(* IEC 61131-3 sources: 2026_Projet_YGO_ExcavatriceDragage/CODE/J_SUPERVISION/_TYPES/2_TRANSLATION, 17 files *)

(* ---- E_TranslationTraceBlockReason.st ---- *)
(* =======================================================================
   🎯 E_TranslationTraceBlockReason — Cause de blocage priorisée translation M3
   ───────────────────────────────────────────────────────────────
   🎯 Rôle : Ordre de priorité de la cause de blocage de la translation M3,
      calculé en PRG_05_Translation et publié via Data.TranslationTrace.
      L'ordre de l'enum EST l'ordre de priorité (valeur croissante = priorité
      décroissante) : la cause la plus grave gagne (PowerCutOff > … > NONE).
   📤 Producteur unique : PRG_05_Translation.
   📥 Consommateur : FB_TroubleshootingView (recopie → GVL_Troubleshooting.S_TraceTranslation).
   🔒 Lecture seule — aucune action de conduite n'en dépend.
   📄 Doc métier : DOC/AF/AF_Partie-14_Fonction_Troubleshooting/FB_TroubleshootingView_v1.2.md
   ======================================================================= *)
{attribute 'qualified_only'}
TYPE E_TranslationTraceBlockReason :
(
    NONE              := 0,   // ✅ Aucun blocage — permis de mouvement effectif
    POWER_CUTOFF      := 1,   // 🧨 Coupure puissance amont (instSafetyTranslationM3.PowerCutOff) — priorité max
    SAFESTOP          := 2,   // 🟧 SafeStop effectif (InputModule OR safety M3)
    SAFETY_FAULT      := 3,   // 🛡️ Défaut safety M3 latched (FB_Safety_Translation.Fault.Error)
    HEIGHT_INTERLOCK  := 4,   // 🚧 Interlock hauteur M1/M2 actif (risque collision)
    DRIVE_UNAVAILABLE := 5,   // 📡 Variateur AC600 injoignable / non opérationnel
    FINAL_INTERLOCK   := 6,   // 🛑 Barrière finale en défaut (frein / redémarrage)
    FAULT             := 7    // ❌ Défaut mouvement M3 latched (FB_Translation.Fault.Error)
);
END_TYPE

(* ---- ST_BypassTranslation.st ---- *)
(* ═══════════════════════════════════════════════════════════════
   ST_BypassTranslation — Bypass maintenance dédiés à Translation M3
   ───────────────────────────────────────────────────────────────
   🔒 Doctrine : actionnable UNIQUEMENT en MAINT_N2, RETAIN, jamais masque
      les autres défauts du même bloc (voir REGISTRE_ACTIONS_Bypass_v1.0 (archive)).
   ═══════════════════════════════════════════════════════════════ *)
TYPE ST_BypassTranslation :
STRUCT
    (* 📡 1. Communication & Systèmes auxiliaires *)
    OperatorComm      : BOOL; (* 📡 Bypass communication esclave CANopen Joystick / heartbeat IHM *)
    DriveComm         : BOOL; (* 📡 Bypass diagnostic esclave EtherCAT AC600 (variateur) *)
    ContactorFeedback : BOOL; (* 🔌 Bypass feedbacks contacteur de frein *)
    PhaseRotation     : BOOL; (* ⚡ Bypass défaut rotation de phases (commun machine) *)
    BrakeThermal      : BOOL; (* 🌡️ Bypass surchauffe thermique frein (commun machine) *)

    (* 🚧 2. Limites physiques et Positionnement *)
    LimitSwitch       : BOOL; (* 🚧 Bypass fins de course physiques avant/arrière *)
    SensorIncoherent  : BOOL; (* 🧭 Bypass incohérence mot capteurs de position *)
    MinHeight         : BOOL; (* : Bypass interlock hauteur mini M1/M2 requise pour translation *)

    (* ⚙️ 3. Sécurité Mécanique (Méca A-B) *)
    MecaA             : BOOL; (* 🔄 Bypass Méca A : mouvement non commandé à l'arrêt *)
    MecaB             : BOOL; (* 🛑 Bypass Méca B : absence confirmation arrêt (frein/contacteurs) *)

    (* 🛡️ 4. Hiérarchie & Restauration *)
    Safety            : BOOL; (* 🛡️ Bypass groupé : tous les bits qui provoquent un PowerCutOff *)
    Process           : BOOL; (* ⚙️ Bypass groupé : tous les bits qui provoquent un SafeStop *)
    Global            : BOOL; (* 🌐 Bypass Global : ignore toutes les sécurités de cet axe *)
    // Flag restauration boot dédié (défaut FALSE non ambigu, contrairement à une valeur métier)
    Initialized       : BOOL := FALSE; (* 🚦 TRUE = bypass restauré depuis GVL_BypassRetain ce boot *)
END_STRUCT
END_TYPE

(* ---- ST_Chain_Translation_Control.st ---- *)
TYPE ST_Chain_Translation_Control :
STRUCT
    Idx401_MotionAllowed         : BOOL; // 1 = Mouvement Translation Autorisé | 0 = Bloqué
    Idx402_SetpointFreq_Hz       : REAL; // [Hz] Consigne Fréquence Calculée
    Idx403_DriveControlWord      : WORD; // Mot de Commande Calculé Variateur AC600
    Idx404_FinalInterlockState   : E_State; // 🛡️ État frontière
    Idx405_FinalInterlockReason  : E_TranslationFinalInterlockReason; // 🛡️ Cause mémorisée
    Idx406_BrakeCommandOpenConfirmed : BOOL; // 🔌 Contacteur/bobine, pas frein mécanique
    Idx407_BrakeTimeoutElapsed   : TIME; // ⏱️ Watchdog 500ms écoulé
END_STRUCT
END_TYPE

(* ---- ST_Chain_Translation_Demandes.st ---- *)
TYPE ST_Chain_Translation_Demandes :
STRUCT
    Idx201_JoyXRaw_ANA           : INT;  // [pts] Bruts Joystick Axe X
    Idx202_JoyXScaled_Pct        : REAL; // [%] Consigne Joystick Axe X (-100% à +100%)
    Idx203_HmiCmd_BtnTremie : BOOL; // 1 = Bouton vers Trémie IHM | 0 = Relâché (ex-Idx203_HmiCmd_BtnFwd)
    Idx204_HmiCmd_BtnMaintenance : BOOL; // 1 = Bouton vers Maintenance IHM | 0 = Relâché (ex-Idx204_HmiCmd_BtnRev)
    Idx205_HmiTargetPosition     : INT;  // Cible Sélectionnée IHM (1=Trémie, 2=P2, 3=P1)
    Idx206_CycleTargetPosition   : INT;  // Cible Sélectionnée par le Cycle Auto
    Idx207_ModeActive            : E_Mode;// Mode courant (MANU_N1, AUTO_N1...)
    Idx208_BypassNetworkActive   : BOOL; // 0 = Comm Variateur OK | 1 = Bypass Réseau Actif ⚠️
    Idx209_ArbitratedSpeed_Pct   : REAL; // [%] Consigne finale Vitesse Translation
END_STRUCT
END_TYPE

(* ---- ST_Chain_Translation_Inputs.st ---- *)
TYPE ST_Chain_Translation_Inputs :
STRUCT
    Idx101_PosTremie_DI          : BOOL; // 1 = Position Trémie Atteinte | 0 = Absent
    Idx102_PosPV_DI              : BOOL; // 1 = Zone Ralentissement PV Atteinte | 0 = Absent
    Idx103_PosP2_DI              : BOOL; // 1 = Position Fosse P2 Atteinte | 0 = Absent
    Idx104_PosP1_DI              : BOOL; // 1 = Position Fosse P1 Atteinte | 0 = Absent
    Idx105_PosMaintenance_DI     : BOOL; // 1 = Position Service Maintenance Atteinte | 0 = Absent
    Idx106_DriveActualFreq_Hz    : REAL; // [Hz] Fréquence Réelle Mesurée Variateur
    Idx107_DriveStatusWord       : WORD; // Mot d'état Brut Variateur AC600
    Idx108_BrakeApplied          : BOOL; // TRUE = frein SERRÉ (NOT BrakeFeedback — IHM garde le sens serré)
    Idx109_DriveThermalOk        : BOOL; // TRUE = thermique moteur/variateur AC600 OK (diagnostic seul)
END_STRUCT
END_TYPE

(* ---- ST_Chain_Translation_Outputs.st ---- *)
TYPE ST_Chain_Translation_Outputs :
STRUCT
    Idx501_CmdDriveControlWord   : WORD; // Mot de Commande Transmis EtherCAT AC600
    Idx502_CmdDriveFreq_Hz       : UINT; // [0.01Hz] Consigne Fréquence Transmise EtherCAT
    Idx503_CmdBrakeRelease_RQ    : BOOL; // 1 = Bobine Frein Translation Alimentée (Ouvert)
END_STRUCT
END_TYPE

(* ---- ST_Chain_Translation_Safety.st ---- *)
TYPE ST_Chain_Translation_Safety :
STRUCT
    Idx301_EmergencyChainClosed  : BOOL; // 1 = Boucle Urgence OK | 0 = Arrêt d'Urgence Appuyé
    Idx302_SafeStopActive        : BOOL; // 0 = Sain (Autorisé) | 1 = Arrêt Rapide Translation
    Idx303_PowerCutOffActive     : BOOL; // 0 = Puissance OK | 1 = Coupure Puissance
    Idx304_LimitSwitchTremieActive  : BOOL; // 0 = Sain | 1 = Fin de Course Extrême Trémie (ex-Idx304_LimitSwitchFwdActive)
    Idx305_LimitSwitchMaintenanceActive : BOOL; // 0 = Sain | 1 = Fin de Course Extrême Maintenance (ex-Idx305_LimitSwitchRevActive)
    Idx306_BypassLimitSwitch     : BOOL; // 0 = Fins de course actives | 1 = Shuntés IHM ⚠️
    Idx307_PositionDecoderIncoherent: BOOL; // 0 = Décodage 5 Capteurs OK | 1 = Incohérence Position
    Idx308_HeightInterlockBlocking: BOOL; // : 0 = M1 ET M2 ≥ hauteur mini (ou bypass) | 1 = Translation bloquée (risque collision)
    (* Défauts safety déchiffrés (bits ErrorId) — visibles individuellement à l'IHM *)
    Idx309_ErrorOperatorComm : BOOL; // bit0 Perte communication opérateur (joystick CAN / heartbeat IHM)
    Idx310_ErrorDriveComm    : BOOL; // bit1 Perte communication EtherCAT variateur
    Idx311_ErrorPhaseRotation: BOOL; // bit2 Mauvaise rotation de phases
    Idx312_ErrorBrakeThermal : BOOL; // bit3 Surchauffe thermique frein commun
    Idx313_ErrorMecaB        : BOOL; // bit4 Absence confirmation arrêt
    Idx314_ErrorMecaA        : BOOL; // bit5 Mouvement non commandé
    Idx315_ErrorLimitSwitch  : BOOL; // bit6 Limite extrême atteinte
    Idx316_ErrorSensorIncoherent: BOOL; // bit7 Mot capteurs position incohérent
    Idx317_ErrorId           : WORD; // Masque brut complet (latch cause) — source d'arbitrage PowerCutOff
    (* Permis directionnels M3 (source unique : FB_Safety_Translation) — TRUE = autorisé, fail-safe *)
    Idx318_EffectivePermitM3_Tremie      : BOOL; // 1 = Translation vers Trémie autorisée | 0 = SENS TRÉMIE BLOQUÉ
    Idx319_EffectivePermitM3_Maintenance : BOOL; // 1 = Translation vers Maintenance/P1 autorisée | 0 = SENS MAINTENANCE BLOQUÉ
END_STRUCT
END_TYPE

(* ---- ST_ChainTranslation.st ---- *)
TYPE ST_ChainTranslation :
STRUCT
    Inputs_100    : ST_Chain_Translation_Inputs;
    Demandes_200  : ST_Chain_Translation_Demandes;
    Safety_300    : ST_Chain_Translation_Safety;
    Control_400   : ST_Chain_Translation_Control;
    Outputs_500   : ST_Chain_Translation_Outputs;
END_STRUCT
END_TYPE

(* ---- ST_HwTranslation.st ---- *)
(* ═══════════════════════════════════════════════════════════════
   🏗️ ST_HwTranslation — Image matérielle brute des entrées Translation M3
   ───────────────────────────────────────────────────────────────
   🎨 Regroupe les signaux physiques d'entrée bruts de la translation M3 (AC600).
   ═══════════════════════════════════════════════════════════════ *)
TYPE ST_HwTranslation :
STRUCT
    M3_PosTremie_DI      : BOOL;         (* Capteur position trémie *)
    M3_PosPV_DI          : BOOL;         (* Capteur position point de vitesse (pré-ralentissement) *)
    M3_PosPVP2_DI        : BOOL;         (* Capteur position P2 / petite vitesse avant P1 *)
    M3_PosP1_DI          : BOOL;         (* Capteur position P1 *)
    M3_PosMaintenance_DI : BOOL;         (* Capteur position maintenance *)
    M3_BrakeIsOpen_DI    : BOOL;         (* Retour frein M3 (1 = ouvert) *)
    M3_ThermalOK_DI      : BOOL;         (* Retour disjoncteur thermique moteur/variateur AC600 (1 = OK) — diagnostic seul, l'AC600 se protège lui-même *)
    M3_StatusWord        : WORD;         (* Status word variateur AC600 *)
    M3_ActualFrequencyHz : UINT;         (* Fréquence réelle variateur AC600 (x100) *)
    AC600_DeviceState    : DEVICE_STATE; (* État device AC600 (GetDeviceState) *)
END_STRUCT
END_TYPE

(* ---- ST_SafetyTranslation.st ---- *)
(* ═══════════════════════════════════════════════════════════════
   🛡️ ST_SafetyTranslation — Diagnostics de sécurité pour la Translation M3
   ───────────────────────────────────────────────────────────────
   🎨 Destiné à l'affichage des défauts de sécurité du translation.
   ═══════════════════════════════════════════════════════════════ *)
TYPE ST_SafetyTranslation :
STRUCT
    Error             : BOOL;    (* 🛡️ Bloc sécurité (Safety) en défaut *)
    ErrorId           : WORD;    (* ❌ Code bitfield du défaut de sécurité (vue LIVE) *)
    LatchedId         : WORD;    (* 🕘 Vue LATCHÉE : ErrorId figé au défaut, effacé au Reset (marqueur [HISTO]) *)
    ErrorOperatorComm : BOOL;    (* 🎮 Perte communication opérateur : joystick CAN ou heartbeat IHM (bit0) *)
    ErrorDriveComm    : BOOL;    (* 📡 Perte communication EtherCAT variateur (bit1) *)
    ErrorPhaseRotation: BOOL;    (* ⚡ Mauvaise rotation de phases électriques (bit2) *)
    ErrorBrakeThermal : BOOL;    (* 🌡️ Surchauffe thermique frein commun (bit3) *)
    ErrorMecaB        : BOOL;    (* 🛑 Absence confirmation arrêt (Méca B - bit4) *)
    ErrorMecaA        : BOOL;    (* 🔄 Mouvement non commandé (Méca A - bit5) *)
    ErrorLimitSwitch  : BOOL;    (* 🚧 Limite extrême Translation atteinte (bit6) *)
    ErrorSensorIncoherent : BOOL; (* 🧭 Mot capteurs M3 incohérent (bit7) *)
    SafeStop          : BOOL;    (* 🛡️ Décélération de sécurité demandée *)
    PowerCutOff       : BOOL;    (* 🧨 Coupure puissance demandée *)
    EffectivePermitM3_Tremie      : BOOL;    (* 🟢 Permis canonique M3 vers Trémie, TRUE = autorisé *)
    EffectivePermitM3_Maintenance : BOOL;    (* 🟢 Permis canonique M3 vers Maintenance/P1, TRUE = autorisé *)
    BlockedBySafety   : BOOL;    (* 🚫 Synthèse globale : translation bloquée par la sécurité *)
    PowerCutOffSafety : BOOL;    (* 🧨 Synthèse sécurités critiques entraînant une coupure puissance *)
    SafeStopSafety    : BOOL;    (* 🛡️ Synthèse défauts entraînant un SafeStop / Rampe rapide *)
END_STRUCT
END_TYPE

(* ---- ST_TraceTranslation.st ---- *)
(* =======================================================================
   ↔️ ST_TraceTranslation — Trace de blocage terrain de la translation M3
   ───────────────────────────────────────────────────────────────
   🎯 Rôle : Publier au technicien « pourquoi la translation M3 ne bouge pas » :
      permis de mouvement effectif, interlock hauteur, source SafeStop/coupure
      et cause de blocage priorisée.
   📤 Producteur unique : PRG_05_Translation (Data.TranslationTrace).
   📥 Consommateur : FB_TroubleshootingView (pure recopie → GVL_Troubleshooting.S_TraceTranslation).
   🔒 Lecture seule — aucun calcul de commande n'en dépend.
   🕒 BlockReasonTimestamp : ms depuis démarrage PLC (TIME()), latched au dernier
      changement de BlockReason (1 scan, mémoire).
   📄 Doc métier : DOC/AF/AF_Partie-14_Fonction_Troubleshooting/FB_TroubleshootingView_v1.2.md
   ======================================================================= *)
TYPE ST_TraceTranslation :
STRUCT
    // Permis de mouvement effectif (agrégat diagnostic : toutes les barrières levées)
    MotionPermitEffective    : BOOL;   // 🟢 Translation réellement autorisée à se déplacer
    // Permis directionnels par sens (reflet exact des permis appliqués au mouvement M3)
    EffectivePermitM3_Tremie      : BOOL;   // 🟢 Permis canonique M3 vers Trémie (reflet lecture seule)
    EffectivePermitM3_Maintenance : BOOL;   // 🟢 Permis canonique M3 vers Maintenance/P1 (reflet lecture seule)
    TremieProcessBlockActive : BOOL;   // 🛑 Approche trémie interdite par process (trémie pleine / grille levée) — recul libre. Motif du permis trémie rouge.
    HeightInterlockBlocking  : BOOL;   // 🚧 Interlock hauteur M1/M2 actif (risque collision)

    // Source de blocage — pour distinguer l'origine
    SafeStopActive           : BOOL;   // 🟧 SafeStop effectif appliqué (M3_SafeStop_Aggregate)
    SafeStopSourceInput      : BOOL;   // 📥 SafeStop issu du module d'entrée (InputModuleFault)
    SafeStopSourceSafety     : BOOL;   // 🛡️ SafeStop issu de FB_Safety_Translation (défaut safety)
    PowerCutOffActive        : BOOL;   // 🧨 Coupure puissance amont active
    DriveOperational         : BOOL;   // 📡 Variateur AC600 opérationnel

    // Barrière finale (frein / redémarrage)
    FinalInterlockError      : BOOL;   // 🛑 Défaut barrière finale (frein / redémarrage)

    // Cause de blocage priorisée + horodatage
    BlockReason              : E_TranslationTraceBlockReason; // 🎯 Cause de blocage prioritaire (ordre de priorité croissant)
    BlockReasonTimestamp     : UDINT;  // 🕒 ms depuis démarrage PLC (TIME()) — dernier changement de BlockReason
END_STRUCT
END_TYPE

(* ---- ST_TranslationCfg.st ---- *)
(* ═══════════════════════════════════════════════════════════════
   ST_TranslationCfg — Configurations et paramètres réglables pour Translation M3
   ───────────────────────────────────────────────────────────────
   🎨 Destiné au paramétrage depuis l'IHM (RETAIN) — même patron que ST_WinchCfg.
   📄 Vitesses de ralentissement d'approche réglables depuis l'IHM (RETAIN), même patron que ST_WinchCfg.
   ═══════════════════════════════════════════════════════════════ *)
TYPE ST_TranslationCfg :
STRUCT
    CfgApproachSpeedTremie_Hz      : REAL := 20.0; (* 🐢 Vitesse réduite d'approche Trémie (Hz), déclenchée par capteur PV, Direction=1 — reglage nominal confirme operateur *)
    CfgApproachSpeedMaintenance_Hz : REAL := 20.0; (* 🐢 Vitesse réduite d'approche Maintenance (Hz), déclenchée par capteur P1, Direction=-1 — reglage nominal confirme operateur *)
    CfgApproachSpeedP1_Hz          : REAL := 20.0; (* 🐢 Vitesse réduite d'approche P1 (Hz), déclenchée par capteur P2, Direction=-1 — reglage nominal confirme operateur *)

    (* Flag restauration boot (défaut FALSE non ambigu) — même patron que ST_WinchCfg *)
    Initialized                    : BOOL := FALSE; (* 🚦 TRUE = config restaurée depuis GVL_PERSISTENT ce boot *)
END_STRUCT
END_TYPE

(* ---- ST_TranslationCmd.st ---- *)
(* ═══════════════════════════════════════════════════════════════
   🎮 ST_TranslationCmd — Commandes IHM pour la Translation M3
   ───────────────────────────────────────────────────────────────
   🎨 Destiné au pilotage de la translation M3 depuis l'IHM.
   📄 : Initialized protège SetFreq_Hz (seul réglage à survivre au reboot),
      sans pont générique pour ne jamais persister BtnTremie/BtnMaintenance.
   ═══════════════════════════════════════════════════════════════ *)
TYPE ST_TranslationCmd :
STRUCT
    SelPositioning     : BOOL;    (* 🎯 TRUE = positionneur sur SelTarget ; FALSE = jog libre *)
    SelTarget          : INT;     (* 🔢 Numéro de la cible de position sélectionnée *)
    BtnTremie         : BOOL;    (* ↔️ Requête marche vers Trémie (ex-BtnFwd), pilotage IHM exclusif *)
    BtnMaintenance    : BOOL;    (* ↔️ Requête marche vers Maintenance (ex-BtnRev), pilotage IHM exclusif *)
    SetFreq_Hz         : REAL;    (* 🎯 Consigne fréquence manuelle [Hz], limitée par PRG_06_Outputs *)
    // 🔀 Switch machine unique : GVL_IHM.Modes.Cmd.TglJoystickMaster (ST_ModesCmd), applicable à M1/M2 ET M3.
    InvertDirection    : BOOL;    (* 🔄 TRUE = inverse Fwd→Maintenance / Rev→Trémie (mise en service) *)
    TglMaintenanceZoneAccess : BOOL; (* : autorisation CONSCIENTE zone Maintenance, EN PLUS de MAINT_N2 (Auth.MaintenanceM3TargetEnable) *)
    TglAllowWinchMoveAtTremie : BOOL; (* T249 : autorisation CONSCIENTE montee/descente treuil couple (WinchSel=0) a la Tremie, EN PLUS de la garde WinchSel=2 forcee (FB_Modes) *)
    Initialized        : BOOL := FALSE; (* 🚦 TRUE = SetFreq_Hz restauré depuis GVL_PERSISTENT ce boot *)
    BtnSetAtP1         : BOOL;    (* 🎯 Forcage position P1 depuis IHM en MAINT_N2 (mise en service) *)
END_STRUCT
END_TYPE

(* ---- ST_TranslationFinalInterlockRequest.st ---- *)
(* ═══════════════════════════════════════════════════════════════
   ↔️ ST_TranslationFinalInterlockRequest — Demande brute vers PDO M3
   ───────────────────────────────────────────────────────────────
   📤 Producteur unique : PRG_05_Translation (VAR_OUTPUT).
   📥 Consommateur unique : PRG_06_Outputs, avant
      FB_TranslationOutputInterlock.
   🔒 Ne contient jamais une commande PDO autorisée.
   PowerCutOff : demande safety M3 (FB_Safety_Translation).
      Consommée par PRG_06_Outputs comme SEULE cause de coupure
      d'Enable (barrière finale). SafeStop est géré en amont
      par FB_Translation (rampe rapide, Enable maintenu, AF06 §5).
   ═══════════════════════════════════════════════════════════════ *)

TYPE ST_TranslationFinalInterlockRequest :
STRUCT
    Enable                       : BOOL;
    Reset                        : BOOL;
    PowerContactorEngaged              : BOOL;
    SafeStop                     : BOOL;
    EffectivePermitM3_Tremie     : BOOL;
    EffectivePermitM3_Maintenance: BOOL;
    PowerCutOff                  : BOOL; // 🧨 Demande coupure puissance (FB_Safety_Translation) — consommée par PRG_06_Outputs (Enable)
    BrakeReleaseRequest          : BOOL;
    BrakeCommandOpenConfirmed    : BOOL; // TRUE = contacteur/bobine desserrage confirmé
    RequestedDriveControlWord    : WORD; // 0=None, 1=Fwd, 2=Rev, 7=Reset AC600
    RequestedDriveFreqHz         : REAL;
    ReqTremieSemantic            : BOOL; // TRUE = mouvement demande vers Tremie, independant de InvertDriveDirection
    ReqMaintenanceSemantic       : BOOL; // TRUE = mouvement demande vers Maintenance/P1, independant de InvertDriveDirection
END_STRUCT
END_TYPE

(* ---- ST_TranslationHMI.st ---- *)
(* ═══════════════════════════════════════════════════════════════
   ↔️ ST_TranslationHMI — Données d'échange IHM pour le Translation M3
   ───────────────────────────────────────────────────────────────
   🎨 Destiné à l'affichage des états, commandes et diagnostics du translation.
   📄 Structuration en Cmd / State / Safety / Bypass / Test —
      doc métier : DOC/AF/AF_Partie-11_Fonction_Translation_v2.3.md
   ═══════════════════════════════════════════════════════════════ *)
TYPE ST_TranslationHMI :
STRUCT
    (* 🎮 Commandes opérateur (manuel / maintenance) *)
    Cmd                     : ST_TranslationCmd;

    (* 🚦 États & diagnostics *)
    State                   : ST_TranslationState;

    (* Configurations et limites — champ Cfg manquait initialement (contrairement à ST_WinchHMI) *)
    Cfg                     : ST_TranslationCfg;

    (* Bypass maintenance *)
    Bypass                  : ST_BypassTranslation;

    (* 🛡️ Sécurité (FB_Safety_Translation) *)
    Safety                  : ST_SafetyTranslation;
END_STRUCT
END_TYPE

(* ---- ST_TranslationInterPrg.st ---- *)
(* ═══════════════════════════════════════════════════════════════
   ↔️ ST_TranslationInterPrg — Bus d'échange inter-PRG produit par PRG_05_Translation
   ───────────────────────────────────────────────────────────────
   🎯 Rôle : Encapsuler la demande finale M3, l'état public TranslationState
      et le diagnostic TranslationSafety publiés par PRG_05_Translation vers
      les consommateurs (PRG_03/06/07).
   📤 Producteur unique : PRG_05_Translation (VAR_OUTPUT Data : ST_TranslationInterPrg).
   📄 Doc : DOC/AF/AF_Partie-11_Fonction_Translation_v2.3.md
   🔌 Architecture : Bus de données typé — encapsulation des échanges inter-PRG.
   ═══════════════════════════════════════════════════════════════ *)

TYPE ST_TranslationInterPrg :
STRUCT
    // === ⚡ Demande finale M3 ===
    TranslationFinalInterlockRequest : ST_TranslationFinalInterlockRequest; // ↔️ Demande finale et interlocks translation M3

    // === 📊 État public translation ===
    TranslationState                 : ST_TranslationState; // 🚦 Etat public translation M3

    // === 🛡️ Sécurité translation ===
    TranslationSafety                : ST_SafetyTranslation; // 🛡️ Diagnostic et securites translation M3

    // === 🎯 Faits decodeur position M3 (produits par PRG_05, AF-02 TBD §8 #5) ===
    M3_SensorWordIncoherent   : BOOL; // ❌ Incoherence detectee mot capteurs M3

    // === ⚙️ États dynamiques & positions stables translation M3 ===
    TranslationBusy           : BOOL; // ⚙️ Translation M3 en mouvement effectif
    TranslationDone           : BOOL; // ✅ Cible translation atteinte et confirmee
    M3_AtTremieStable         : BOOL; // 🎯 M3 positionne stable a la Tremie
    M3_AtP1Stable             : BOOL; // 🎯 M3 positionne stable au Point 1
    M3_AtMaintenanceStable    : BOOL; // 🎯 M3 positionne stable en zone Maintenance
    M3_AtWorkPositionStable   : BOOL; // 🎯 M3 arrete a une position de travail (P1 ou Maintenance) — STATIQUE (mot capteurs), vrai des le boot sans franchissement. Consomme par le verrou descente treuil T249-A.

    // === 🕵️ Trace de blocage terrain (consommée FB_TroubleshootingView) ===
    TranslationTrace             : ST_TraceTranslation; // 🕵️ Trace blocage translation M3 (cause priorisée + horodatage)
END_STRUCT
END_TYPE

(* ---- ST_TranslationState.st ---- *)
(* ═══════════════════════════════════════════════════════════════
   🚦 ST_TranslationState — États et retours IHM pour la Translation M3
   ───────────────────────────────────────────────────────────────
   🎨 Destiné à l'affichage des retours et mesures de la translation M3.
   ═══════════════════════════════════════════════════════════════ *)
TYPE ST_TranslationState :
STRUCT
    (* 🚦 États & diagnostics FB_Translation *)
    FBState                 : E_State; (* 🤖 État de l'automate interne (FB_Translation) *)
    AxisBlockReason         : E_TranslationTraceBlockReason; (* 🧩 Cause prioritaire de blocage (miroir de TranslationTrace.BlockReason) *)
    Ready                   : BOOL;    (* 🟢 Translation prêt à fonctionner *)
    Busy                    : BOOL;    (* ⚙️ Mouvement en cours *)
    Done                    : BOOL;    (* ✅ Mouvement terminé avec succès *)
    Error                   : BOOL;    (* Translation en défaut *)
    ErrorId                 : WORD;    (* ❌ Code du défaut actif *)
    BrakeCmd                : BOOL;    (* 🔓 Commande de desserrage du frein (lecture seule, TRUE = desserré) *)
    BrakeFeedback           : BOOL;    (* 🔌 Retour physique direct : TRUE = frein OUVERT (desserré) *)
    PositionSensorTarget    : BOOL;    (* 🎯 Capteur de détection de la position cible atteint *)
    PositionReached         : BOOL;    (* ✅ Positionneur : cible sélectionnée atteinte (non mémorisé) *)
    DriveActualFreq_Hz      : REAL;    (* 📈 Fréquence de sortie réelle du variateur (Hz) *)
    DriveControlWord        : WORD;    (* ⚙️ Mot de commande AC600 réellement appliqué *)
    DriveFreqCmd_Hz         : REAL;    (* 🎯 Commande fréquence réellement appliquée *)
    ActiveTremie            : BOOL;    (* ↔️ Commande active vers Trémie *)
    ActiveMaintenance       : BOOL;    (* ↔️ Commande active vers Maintenance *)
    SpeedCmd_Pct            : REAL;    (* 📊 Commande active après arbitrage (0.0 à 100.0 %) *)
    FinalInterlockState     : E_State; (* 🛡️ État final lecture seule *)
    FinalInterlockReason    : E_TranslationFinalInterlockReason; (* 🛡️ Cause finale mémorisée *)
    FinalInterlockError     : BOOL;    (* 🛡️ Défaut final mémorisé *)
    FinalInterlockErrorId   : WORD;    (* 🛡️ Bitfield final *)
    BrakeCommandOpenConfirmed : BOOL;  (* 🔌 Contacteur/bobine desserrage confirmé, pas frein mécanique *)
    FinalBrakeTimeoutElapsed : TIME;   (* ⏱️ Écoulé watchdog 500ms *)

    (* 🔌 Diagnostic variateur EtherCAT (décodé — pas de bit-masking côté IHM) *)
    DriveCommReady          : BOOL;    (* 📡 Variateur M3 : communication prête (StatusWord bit7) *)
    DrivePowerReady         : BOOL;    (* ⚡ Variateur M3 : puissance prête (StatusWord bit0) *)

    (* 📍 Mot capteurs et positions Translation M3 *)
    PositionTremie          : BOOL;
    PositionPV              : BOOL;
    PositionP2              : BOOL;
    PositionP1              : BOOL;
    PositionMaintenance     : BOOL;
    (* : mot EXACT — front franc arrivée/cible (voir PositionXxx ci-dessus = cumulatif zone, réservé ralentissement) *)
    AtTremie                : BOOL;    (* jeton "dernier capteur franchi" (front + libération sur mouvement confirmé) — logique de positionnement *)
    AtPV                    : BOOL;
    AtP2                    : BOOL;
    AtP1                    : BOOL;
    AtMaintenance           : BOOL;
    M3StatusText            : STRING(80);  (* T249-B : texte statut position M3 (INFO, lecture seule) — jeton "at position" sur front capteur sinon zone SensorsWord. Ex "M3 a P1 -> Maintenance", "M3 entre P2 et P1" *)
    EstimatedPosM3_M        : REAL;    (* 📏 Position continue estimée en mètres (0.0 m Maint -> +X m Trémie) — persistante, survit reboot *)
    SensorsWord             : BYTE;    (* bit4=Trémie, bit3=PV, bit2=P2, bit1=P1, bit0=Maintenance *)
    SensorWordIncoherent    : BOOL;
    LimitSwitchTremie       : BOOL;    (* 🚧 Fin de course extrême Trémie (ex-LimitSwitchFwd) *)
    LimitSwitchMaintenance  : BOOL;    (* 🚧 Fin de course extrême Maintenance (ex-LimitSwitchRev) *)
    DriveThermalOk          : BOOL;    (* Retour disjoncteur thermique moteur/variateur AC600 — diagnostic seul, l'AC600 se protège lui-même *)
    MaintenanceTargetEnable : BOOL;    (* 🔓 TRUE = Autorise le déplacement vers la cible 4 (Maintenance) ; actif uniquement en mode MAINT_N2 *)
    SimulationModeActive    : BOOL;
    HeightInterlockBlocking : BOOL;    (* : TRUE = translation bloquée, M1 ou M2 sous la hauteur mini requise *)

    (* 📏 T301 — Odométrie M3 : gain actif + mesure PROPOSÉE P2 <-> PV (jamais appliquée, recopie manuelle) *)
    OdometryGainActive            : REAL;   (* Gain consommé par l'estimateur, m/(Hz.s) *)
    OdometryCalibValid            : BOOL;   (* TRUE = gain calculé depuis le réglage Calib* (défaut 2,0 s compris) ; FALSE = gain de repli *)
    OdometryMeasureActive         : BOOL;   (* Mesure P2 <-> PV en cours *)
    OdometryMeasuredTime_S        : REAL;   (* Dernier temps mesuré P2 <-> PV (s) -> à recopier dans _TranslationCalibTimeP2PV_S *)
    OdometryMeasuredFreqAvg_Hz    : REAL;   (* Fréquence moyenne de la mesure (Hz) -> à recopier dans _TranslationCalibFreq_Hz *)
    OdometryMeasuredFreqSpread_Hz : REAL;   (* Écart max - min de fréquence : petit = vitesse constante, mesure fiable *)
    OdometryMeasuredGain          : REAL;   (* Gain qui résulterait de la mesure, m/(Hz.s) *)
    OdometryMeasureCount          : UDINT;  (* Nombre de mesures abouties depuis le démarrage *)
END_STRUCT
END_TYPE
